// TwinCAT 3 PLC project Tutorial_PLC
// ProgramVersion: 3.1.4024.0
// libraries:
//   Swa_PackML, * (SoftWear Automation Inc)
//   Tc2_MC2, * (Beckhoff Automation GmbH)
//   Tc2_Standard, * (Beckhoff Automation GmbH)
//   Tc2_System, * (Beckhoff Automation GmbH)
//   Tc3_Module, * (Beckhoff Automation GmbH)
// project tree:
//   / GlobalTextList.TcGTLO, PlcTask.TcTTO, Visualization Manager.TcVMO (not stored), VISU_TASK.TcTTO
//   GVLs/ TT_GIO.TcGVL
//   Modules/CM_ControlModule/ CM_ControlModule.TcPOU
//   Modules/CM_ControlModule/Enums/ E_CmControlModuleCmd.TcDUT, E_CmControlModuleState.TcDUT
//   Modules/CM_ControlModule/Interfaces/ I_CmControlModule.TcIO
//   Modules/CM_ControlModule/Sequences/ SEQ_ModuleSequence.TcPOU
//   Modules/CM_ControlModule/Structs/ ST_ControlModuleDevList.TcDUT
//   Modules/UM_Tutorial/Enums/ E_UmTutorialCmd.TcDUT, E_UmTutorialState.TcDUT
//   Modules/UM_Tutorial/Interfaces/ I_UmTutorial.TcIO
//   Modules/UM_Tutorial/ UM_Tutorial.TcPOU
//   POUs/ MAIN.TcPOU
//   VISUs/ Visualization.TcVIS
// real-time tasks:
//   TASK PlcTask: cycle T#10ms, priority 20, ADS port 350
//   TASK VISU_TASK: cycle T#200000us, priority 30, ADS port 351
// motion (NC):
//   TASK NC-Task 1 SAF: cycle T#2ms, priority 4, ADS port 501
//   TASK NC-Task 1 SVB: cycle T#10ms, priority 8, ADS port 511
//   AXIS Tutorial Axis (id 1)
//     OtherSettings: AllowMotionCmdToSlave=true
//     encoder EncType=1
//     drive DrvType=5
//       Analog: TorqueSetpointScale=10, ScaleFactorActTorque=0.1
//       TimeComp: TaskDelayCycles=1
//     controller CtrType=1
//       CtrPara: PriorControlFactor=1
//         Observer: BandWidth=20
// I/O:
//   DEVICE LaptopPort (EtherCAT), AmsNetId 10.0.2.15.2.1
//     Rack_01 (EK1101) [EK1100 EtherCAT Coupler (2A E-Bus)]
//       Rack_01_S01 (EL1008) [EL1008 8Ch. Dig. Input 24V, 3ms]
//       Rack_01_S02 (EL9186) [EL9186 Potential Connection, 8 x 24V]
//       Rack_01_S03 (EL9187) [EL9187 Potential Connection, 8 x Ground]
//       Rack_01_S04 (EL2008) [EL2008 8Ch. Dig. Output 24V, 0.5A]
//       Rack_01_S05 (EL7211-9014) [EL7211-9014 1Ch. MDP742 Servo motor output stage with OCT (50V, 4.5A RMS) and STO input]
//       Rack_01_S06 (EL6910) [EL6910, TwinSAFE PLC]
//       Rack_01_S07 (EL2911) [EL2911, Potential supply terminal (10 A) with 4 Ch. Safety Inputs, TwinSAFE]
//         modules: Module 1 (FSOE), Module 2 (FSOUT), Module 3 (DEVICEIO), Module 4 (FSLOGIC)
// variable links:
//   Tutorial_PLC/Tutorial_PLC Instance <-> LaptopPort (EtherCAT)/Rack_01 (EK1101)/Rack_01_S01 (EL1008)
//     PlcTask Inputs/TT_GIO.I_PB_MOMENTARY <-> Channel 2/Input
//     PlcTask Inputs/TT_GIO.I_PB_SAFETY_RESET <-> Channel 1/Input
//     PlcTask Inputs/TT_GIO.I_PX_CYL_EXAMPLE_E <-> Channel 3/Input
//     PlcTask Inputs/TT_GIO.I_PX_CYL_EXAMPLE_R <-> Channel 4/Input
//     PlcTask Inputs/TT_GIO.I_R01_S01_I_BIT_05 <-> Channel 5/Input
//     PlcTask Inputs/TT_GIO.I_R01_S01_I_BIT_06 <-> Channel 6/Input
//     PlcTask Inputs/TT_GIO.I_R01_S01_I_BIT_07 <-> Channel 7/Input
//     PlcTask Inputs/TT_GIO.I_R01_S01_I_BIT_08 <-> Channel 8/Input
//   Tutorial_PLC/Tutorial_PLC Instance <-> LaptopPort (EtherCAT)/Rack_01 (EK1101)/Rack_01_S04 (EL2008)
//     PlcTask Outputs/TT_GIO.O_DO_SIGNAL_PL <-> Channel 7/Output
//     PlcTask Outputs/TT_GIO.O_R01_S04_O_BIT_01 <-> Channel 1/Output
//     PlcTask Outputs/TT_GIO.O_R01_S04_O_BIT_02 <-> Channel 2/Output
//     PlcTask Outputs/TT_GIO.O_R01_S04_O_BIT_03 <-> Channel 3/Output
//     PlcTask Outputs/TT_GIO.O_R01_S04_O_BIT_04 <-> Channel 4/Output
//     PlcTask Outputs/TT_GIO.O_R01_S04_O_BIT_05 <-> Channel 5/Output
//     PlcTask Outputs/TT_GIO.O_R01_S04_O_BIT_06 <-> Channel 6/Output
//     PlcTask Outputs/TT_GIO.O_SV_CYL_EXAMPLE_E <-> Channel 8/Output
//   Tutorial_PLC/Tutorial_PLC Instance <-> NC-Task 1 SAF/Axes/Tutorial Axis
//     PlcTask Inputs/TT_GIO.AX_TUTORIAL.NcToPlc <-> Outputs/ToPlc
//     PlcTask Outputs/TT_GIO.AX_TUTORIAL.PlcToNc <-> Inputs/FromPlc

CONFIGURATION Tutorial_PLC
    RESOURCE PLC ON TwinCAT3
        TASK PlcTask(INTERVAL := T#10ms, PRIORITY := 20);
        TASK VISU_TASK(INTERVAL := T#200000us, PRIORITY := 30);
        PROGRAM MAIN WITH PlcTask : MAIN;
        PROGRAM VisuElems_Visu_Prg WITH VISU_TASK : VisuElems.Visu_Prg;
    END_RESOURCE
END_CONFIGURATION

// ---- Modules/CM_ControlModule/Enums/E_CmControlModuleCmd.TcDUT
{attribute 'qualified_only'}
{attribute 'strict'}
TYPE E_CmControlModuleCmd :
(
	NoCmd
);
END_TYPE

// ---- Modules/CM_ControlModule/Enums/E_CmControlModuleState.TcDUT
{attribute 'qualified_only'}
{attribute 'strict'}
TYPE E_CmControlModuleState :
(
	NoCmd
);
END_TYPE

// ---- Modules/CM_ControlModule/Structs/ST_ControlModuleDevList.TcDUT
TYPE ST_ControlModuleDevList :
STRUCT
	DiMomentaryPb	: I_DevDigitalIn;
	CylExample		: I_DevCylinder;
	DoSignalPl		: I_DevDigitalOut;
END_STRUCT
END_TYPE

// ---- Modules/UM_Tutorial/Enums/E_UmTutorialCmd.TcDUT
{attribute 'qualified_only'}
{attribute 'strict'}
TYPE E_UmTutorialCmd :
(
	NoCmd
);
END_TYPE

// ---- Modules/UM_Tutorial/Enums/E_UmTutorialState.TcDUT
{attribute 'qualified_only'}
{attribute 'strict'}
TYPE E_UmTutorialState :
(
	NoCmd
);
END_TYPE

// ---- GVLs/TT_GIO.TcGVL
{attribute 'qualified_only'}
VAR_GLOBAL
	// TwinSAFE
	Safety	: TwinSAFE;
	// AXIS IO
	//SLICE AXIS
	{attribute 'TcNcAxis' := 'Tutorial Axis'}
	AX_TUTORIAL				: AXIS_REF;  //EL7211-9014 R01 S05
	// SLICE IO
	// TUTORIAL R01 EL1008 SLOT 01
    {attribute 'TcLinkTo' := 'TIID^LaptopPort (EtherCAT)^Rack_01 (EK1101)^Rack_01_S01 (EL1008)^Channel 1^Input'}
	I_PB_SAFETY_RESET		AT %I* : BOOL;
	{attribute 'TcLinkTo' := 'TIID^LaptopPort (EtherCAT)^Rack_01 (EK1101)^Rack_01_S01 (EL1008)^Channel 2^Input'}
	I_PB_MOMENTARY		AT %I* : BOOL;
	{attribute 'TcLinkTo' := 'TIID^LaptopPort (EtherCAT)^Rack_01 (EK1101)^Rack_01_S01 (EL1008)^Channel 3^Input'}
	I_PX_CYL_EXAMPLE_E		AT %I* : BOOL;
	{attribute 'TcLinkTo' := 'TIID^LaptopPort (EtherCAT)^Rack_01 (EK1101)^Rack_01_S01 (EL1008)^Channel 4^Input'}
	I_PX_CYL_EXAMPLE_R		AT %I* : BOOL;
	{attribute 'TcLinkTo' := 'TIID^LaptopPort (EtherCAT)^Rack_01 (EK1101)^Rack_01_S01 (EL1008)^Channel 5^Input'}
	I_R01_S01_I_BIT_05		AT %I* : BOOL;
	{attribute 'TcLinkTo' := 'TIID^LaptopPort (EtherCAT)^Rack_01 (EK1101)^Rack_01_S01 (EL1008)^Channel 6^Input'}
	I_R01_S01_I_BIT_06		AT %I* : BOOL;
	{attribute 'TcLinkTo' := 'TIID^LaptopPort (EtherCAT)^Rack_01 (EK1101)^Rack_01_S01 (EL1008)^Channel 7^Input'}
	I_R01_S01_I_BIT_07		AT %I* : BOOL;
	{attribute 'TcLinkTo' := 'TIID^LaptopPort (EtherCAT)^Rack_01 (EK1101)^Rack_01_S01 (EL1008)^Channel 8^Input'}
	I_R01_S01_I_BIT_08		AT %I* : BOOL;
	// TUTORIAL R01 EL2008 SLOT 04
	{attribute 'TcLinkTo' := 'TIID^LaptopPort (EtherCAT)^Rack_01 (EK1101)^Rack_01_S04 (EL2008)^Channel 1^Output'}
    O_R01_S04_O_BIT_01		AT %Q* : BOOL;
	{attribute 'TcLinkTo' := 'TIID^LaptopPort (EtherCAT)^Rack_01 (EK1101)^Rack_01_S04 (EL2008)^Channel 2^Output'}
    O_R01_S04_O_BIT_02		AT %Q* : BOOL;
	{attribute 'TcLinkTo' := 'TIID^LaptopPort (EtherCAT)^Rack_01 (EK1101)^Rack_01_S04 (EL2008)^Channel 3^Output'}
    O_R01_S04_O_BIT_03		AT %Q* : BOOL;
	{attribute 'TcLinkTo' := 'TIID^LaptopPort (EtherCAT)^Rack_01 (EK1101)^Rack_01_S04 (EL2008)^Channel 4^Output'}
    O_R01_S04_O_BIT_04		AT %Q* : BOOL;
	{attribute 'TcLinkTo' := 'TIID^LaptopPort (EtherCAT)^Rack_01 (EK1101)^Rack_01_S04 (EL2008)^Channel 5^Output'}
    O_R01_S04_O_BIT_05		AT %Q* : BOOL;
	{attribute 'TcLinkTo' := 'TIID^LaptopPort (EtherCAT)^Rack_01 (EK1101)^Rack_01_S04 (EL2008)^Channel 6^Output'}
    O_R01_S04_O_BIT_06		AT %Q* : BOOL;
	{attribute 'TcLinkTo' := 'TIID^LaptopPort (EtherCAT)^Rack_01 (EK1101)^Rack_01_S04 (EL2008)^Channel 7^Output'}
    O_DO_SIGNAL_PL		AT %Q* : BOOL;
	{attribute 'TcLinkTo' := 'TIID^LaptopPort (EtherCAT)^Rack_01 (EK1101)^Rack_01_S04 (EL2008)^Channel 8^Output'}
    O_SV_CYL_EXAMPLE_E		AT %Q* : BOOL;
END_VAR

// ---- Modules/CM_ControlModule/Interfaces/I_CmControlModule.TcIO
INTERFACE I_CmControlModule EXTENDS I_PmlObject

END_INTERFACE

// ---- Modules/UM_Tutorial/Interfaces/I_UmTutorial.TcIO
INTERFACE I_UmTutorial EXTENDS I_PmlObject

END_INTERFACE

// ---- POUs/MAIN.TcPOU
PROGRAM MAIN
VAR
	Machine : UM_Tutorial := (Description := ' Tutorial Project ',
							UseGenericVISU := TRUE);
	DownloadBit : BOOL := TRUE;
END_VAR

TT_GIO.Safety(Reset_Trigger := Machine.PbReset.Actuate);
TT_GIO.Safety.In.EStop_OK := TRUE;
TT_GIO.Safety.In.EStop_STO := TRUE;

Machine(SafetyBlock := TT_GIO.Safety);

END_PROGRAM

// ---- Modules/UM_Tutorial/UM_Tutorial.TcPOU
FUNCTION_BLOCK FINAL UM_Tutorial EXTENDS PML_UnitMachine IMPLEMENTS I_UmTutorial

VAR
	// Tags trailing properties


	// PB Instance Declaration


	// Sequence Instance Declaration


	// Module/Device Instance Declaration
	
	DiResetPb			: DEV_DigitalIn	:= (Description := 'Reset PB'); //Machine Reset Pushbutton Attach to the Unit Machine for uses beyond ESTOP reset
	DiMomentaryPb		: DEV_DigitalIn	:= (Description := 'Momentary PB');
	CylExample			: DEV_Cylinder := (Description := 'Example Cyl', ValveType := E_ValveType.Five2SingleNR, ViewedAsEngDiseng := FALSE, RetractIsEngaged := FALSE);
	DoSignalPl			: DEV_DigitalOut := (Description := 'Signal Pilot Light');
    cmModule			: CM_ControlModule	:= (Description	:= 'Control Module',
											UseGenericVisu	:= TRUE,
											HasParams := FALSE,
											HasStatus := FALSE);	
	//DevLists
	ModuleDevList	: ST_ControlModuleDevList := (DiMomentaryPb	:= DiMomentaryPb,
													CylExample		:= CylExample,
													DoSignalPl		:= DoSignalPl);
											
	// Other local variables
	cmd	: E_UmTutorialCmd;

END_VAR

// Call Pushbutton FBs (or Update command)


// Evaluate commands to drive states, run methods of devices (ax.MoveAbs), run seq etc.
StateTransitionLogic();

// Call Sequence FBs




// Call Module/Device FBs
SUPER^(); // Basically a module. Call other modules below this.
DiResetPb();
DiMomentaryPb();
CylExample();
DoSignalPl();
cmModule(DevList := ModuleDevList);

// Reset cmd at end of FB Scan
cmd := E_UmTutorialCmd.NoCmd;

PROPERTY Empty : BOOL
END_PROPERTY

METHOD PRIVATE InitAlarms : BOOL
END_METHOD

METHOD MapInputs : BOOL
VAR_INPUT
END_VAR
END_METHOD

METHOD MapOutputs : BOOL
VAR_INPUT
END_VAR
END_METHOD

METHOD PRIVATE RaiseAlarm : BOOL
VAR_INPUT
	AlarmId : UDINT;
END_VAR
CASE AlarmId OF
0:
	;
END_CASE
END_METHOD

METHOD PROTECTED RunPmlExecute
// Add custom implementation
CASE CurrentPmlMode OF
	E_PmlMode.Production:
		//

	E_PmlMode.SemiAuto:
		//

	E_PmlMode.Manual:
		//

END_CASE
END_METHOD

METHOD PROTECTED SetDependency
// Attach Sequences


// Attach Modules/Devices
Attach(DiResetPb);
Attach(cmModule);

SUPER^.SetDependency(); // Call at the end, after all of the attach
END_METHOD

METHOD PRIVATE StateTransitionLogic
END_METHOD

END_FUNCTION_BLOCK

// ---- Modules/CM_ControlModule/CM_ControlModule.TcPOU
FUNCTION_BLOCK FINAL CM_ControlModule EXTENDS PML_Module IMPLEMENTS I_CmControlModule
VAR_IN_OUT
    DevList : ST_ControlModuleDevList;
END_VAR
VAR
	// Tags trailing properties


	// PB Instance Declaration


	// Sequence Instance Declaration
	seqModuleSequence	: SEQ_ModuleSequence := (Description := 'Module Sequence', _enableHmiStart := TRUE, _enableSfcTipCtrl := FALSE);

	// Module/Device Instance Declaration

	// Other local variables
	cmd	: E_CmControlModuleCmd;

END_VAR

// Call Pushbutton FBs (or Update command)


// Evaluate commands to drive states, run methods of devices (ax.MoveAbs), run seq etc.
StateTransitionLogic();

// Call Sequence FBs
// Call Sequence FBs
seqModuleSequence(DevList := THIS^.DevList);

// Call Module/Device FBs
SUPER^(); // Basically a module. Call other modules below this.


// Reset cmd at end of FB Scan
cmd := E_CmControlModuleCmd.NoCmd;

METHOD PRIVATE InitAlarms : BOOL
END_METHOD

METHOD PRIVATE RaiseAlarm : BOOL
VAR_INPUT
	AlarmId : UDINT;
END_VAR
CASE AlarmId OF
0:
	;
END_CASE
END_METHOD

METHOD PROTECTED RunPmlExecute
// Add custom implementation
CASE CurrentPmlMode OF
	E_PmlMode.Production:
		//

	E_PmlMode.SemiAuto:
		//

	E_PmlMode.Manual:
		//

END_CASE
END_METHOD

METHOD PROTECTED SetDependency
// Attach Sequences
Attach(seqModuleSequence);

// Attach Modules/Devices

// The warning can be disabled here as the user is aware of the risk that the reference may not be valid by checking its validity
{warning disable C0371}

// Checking the VAR_IN_OUT reference, leave the current method in case of invalid reference
IF NOT __ISVALIDREF(DevList) THEN
     RETURN;
END_IF

// Access to VAR_IN_OUT reference (only if the reference was confirmed as valid before)
AttachDevList(ListPointer := ADR(DevList), ListSize := SIZEOF(DevList));

// The warning may be restored at the end of the access area
{warning restore C0371}
SUPER^.SetDependency(); // Call at the end, after all of the attach
END_METHOD

METHOD PRIVATE StateTransitionLogic
END_METHOD

END_FUNCTION_BLOCK

// ---- Modules/CM_ControlModule/Sequences/SEQ_ModuleSequence.TcPOU
FUNCTION_BLOCK FINAL SEQ_ModuleSequence EXTENDS GEN_Sequence
VAR_IN_OUT
    DevList : ST_ControlModuleDevList;
END_VAR
VAR
END_VAR

SUPER^();

METHOD PRIVATE InitAlarms : BOOL
END_METHOD

METHOD PRIVATE RaiseAlarm : BOOL
VAR_INPUT
	AlarmId : UDINT;
END_VAR
CASE AlarmId OF
0:
	;
END_CASE
END_METHOD

METHOD PROTECTED RunSteps
Steps();
END_METHOD

ACTION Steps:
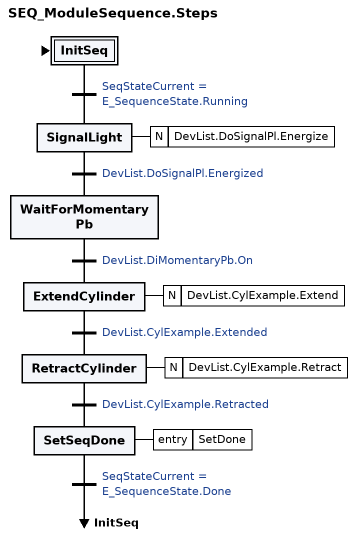
INITIAL_STEP InitSeq:
END_STEP
TRANSITION FROM InitSeq TO SignalLight
    := SeqStateCurrent = E_SequenceState.Running;
END_TRANSITION
STEP SignalLight:
    DevList.DoSignalPl.Energize(N);
END_STEP
TRANSITION FROM SignalLight TO WaitForMomentaryPb
    := DevList.DoSignalPl.Energized;
END_TRANSITION
STEP WaitForMomentaryPb:
END_STEP
TRANSITION FROM WaitForMomentaryPb TO ExtendCylinder
    := DevList.DiMomentaryPb.On;
END_TRANSITION
STEP ExtendCylinder:
    DevList.CylExample.Extend(N);
END_STEP
TRANSITION FROM ExtendCylinder TO RetractCylinder
    := DevList.CylExample.Extended;
END_TRANSITION
STEP RetractCylinder:
    DevList.CylExample.Retract(N);
END_STEP
TRANSITION FROM RetractCylinder TO SetSeqDone
    := DevList.CylExample.Retracted;
END_TRANSITION
STEP SetSeqDone:
    SetDone(P1);  // entry action
END_STEP
TRANSITION FROM SetSeqDone TO InitSeq
    := SeqStateCurrent = E_SequenceState.Done;
END_TRANSITION
END_ACTION

END_FUNCTION_BLOCK

// ---- VISUs/Visualization.TcVIS
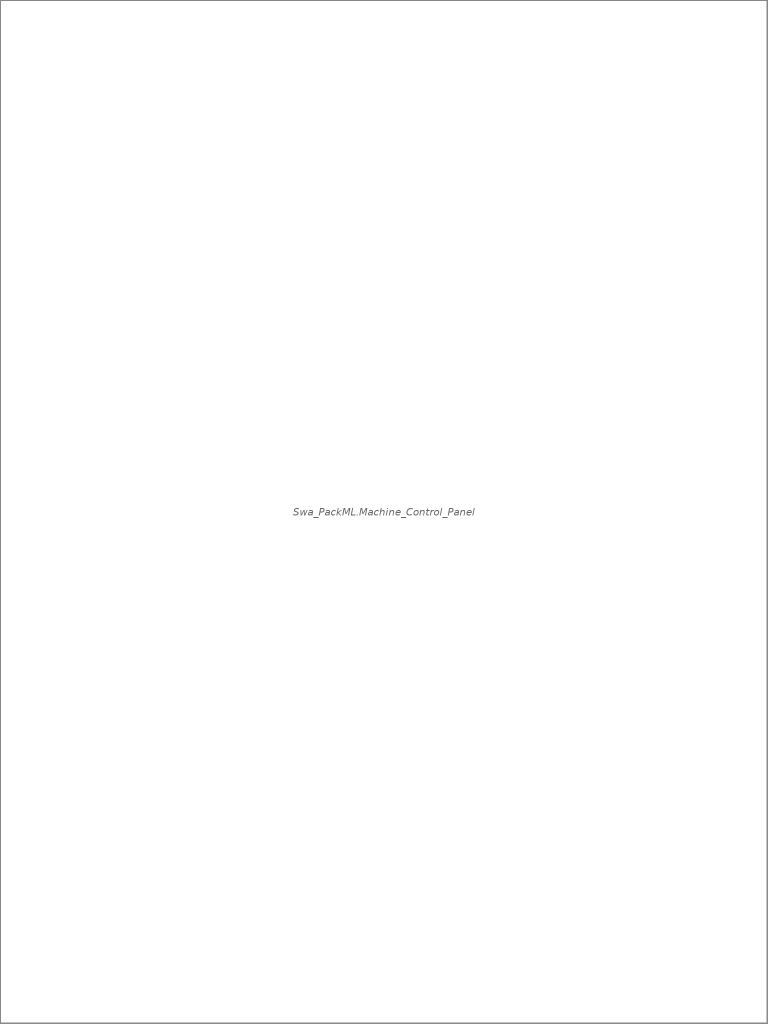
VISUALIZATION Visualization  // 768x1024
    Frame (0,0 768x1024)
        shows Swa_PackML.Machine_Control_Panel(AlarmAdmin := MAIN.Machine.alarmAdmin, ModuleSelector := MAIN.Machine.moduleSelector)
END_VISUALIZATION
